(* Logix 5000 project; controller TFF vendor 1 type 14 code 107 rev 33.11; software revision 33.04; part 17 of 38 *)
(* tags used below, declared in another part *)
   PCV101_AutoMaxRate : REAL;   // PCV101 Maximum Rate in Auto Mode
   PCV101_ManualMaxRate : REAL;   // PCV101 Maximum Rate in Manual mode
   PCV101_Max_CV : REAL;   // Max CV for PCV101
   ControlLoop : ControlLoop[20];   // Control Loop Array
   ControlLoop_PCV101 : ALIAS FOR ControlLoop[3];
   ControlLoop_PCV101_5ms : ALIAS FOR ControlLoop[4];
   ControlLoop_PCV101Alarm : ALIAS FOR AlarmDeviation[3];
   ControlLoop_PCV201 : ALIAS FOR ControlLoop[5];
   ControlLoop_PCV201_5ms : ALIAS FOR ControlLoop[6];
   ControlLoop_PCV201_RAMP_OUT : REAL;   // Ramp Output
   PCV101 : ALIAS FOR AnalogPoint[3];
   PCV101_AO : ALIAS FOR AnalogOutput[3];
   PCV101_Control : PCV_Control;   // PCV101 Control UDT
   PCV101_CVTune : CVTune;
   PCV101_PID : PCV;   // PCV101 PID Management
   PCV201 : ALIAS FOR AnalogPoint[4];
   PCV201_Control : PCV_Control;   // PCV201 Control UDT
   PCV201_PID : PCV;   // PCV201 PID Management
   Rack_Murr_Node1_TFF20 : IO_Station;   // Status of Node 1 TFF20
   Rack_Murr_Node1_TFF40 : IO_Station;   // Status of Node 1 TFF40
   Rack_Murr_Node1_TFF80 : IO_Station;   // Status of Node 1 TFF80
   RawAnalogInputArray : INT[50];   // Array of analog input raw
   SysControl : SysControl;   // General system status and command
   ThisSystem : SystemType;
   TMP : ALIAS FOR AnalogPoint[41];
   Valve : Valve[100];   // Valve Array
(* MainProgram5ms, continued *)

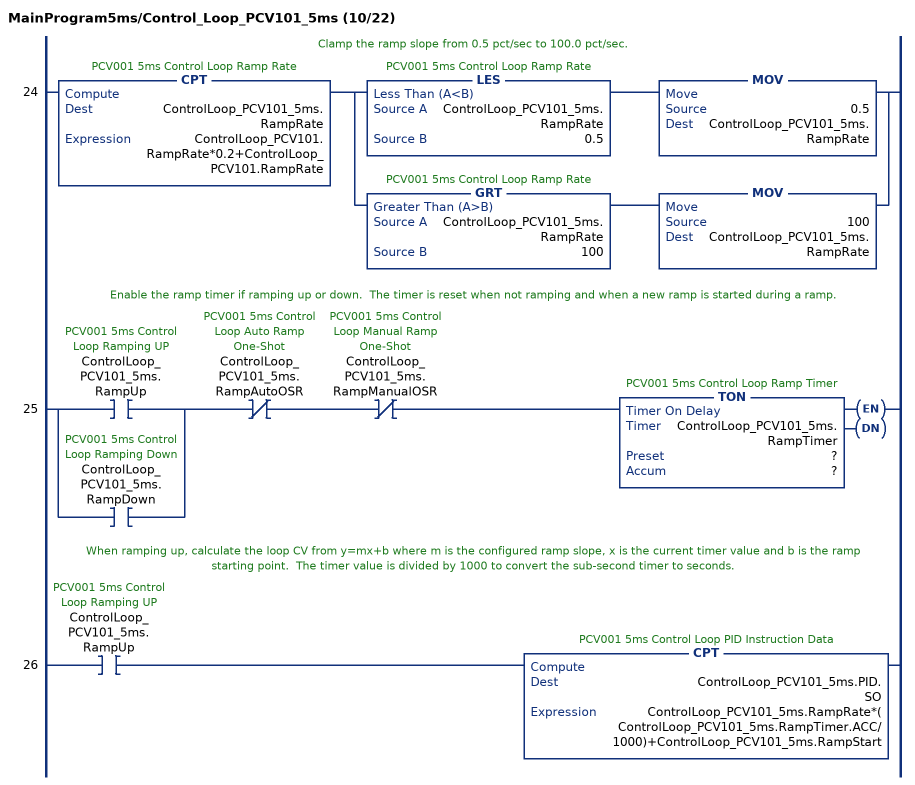
   [picture p62: MainProgram5ms/Control_Loop_PCV101_5ms rungs 24-26]
   // Clamp the ramp slope from 0.5 pct/sec to 100.0 pct/sec.
   24: CPT(ControlLoop_PCV101_5ms.RampRate,ControlLoop_PCV101.RampRate*0.2+ControlLoop_PCV101.RampRate)[LES(ControlLoop_PCV101_5ms.RampRate,0.5) MOV(0.5,ControlLoop_PCV101_5ms.RampRate) ,GRT(ControlLoop_PCV101_5ms.RampRate,100) MOV(100,ControlLoop_PCV101_5ms.RampRate) ];
   // Enable the ramp timer if ramping up or down.  The timer is reset when not ramping and when a new ramp is started during a ramp.
   25: [XIC(ControlLoop_PCV101_5ms.RampUp) ,XIC(ControlLoop_PCV101_5ms.RampDown) ]XIO(ControlLoop_PCV101_5ms.RampAutoOSR)XIO(ControlLoop_PCV101_5ms.RampManualOSR)TON(ControlLoop_PCV101_5ms.RampTimer,?,?);
   // When ramping up, calculate the loop CV from y=mx+b where m is the configured ramp slope, x is the current timer value and b is the ramp starting point.  The timer value is divided by 1000 to convert the sub-second timer to seconds.
   26: XIC(ControlLoop_PCV101_5ms.RampUp)CPT(ControlLoop_PCV101_5ms.PID.SO,ControlLoop_PCV101_5ms.RampRate*(ControlLoop_PCV101_5ms.RampTimer.ACC/1000)+ControlLoop_PCV101_5ms.RampStart);
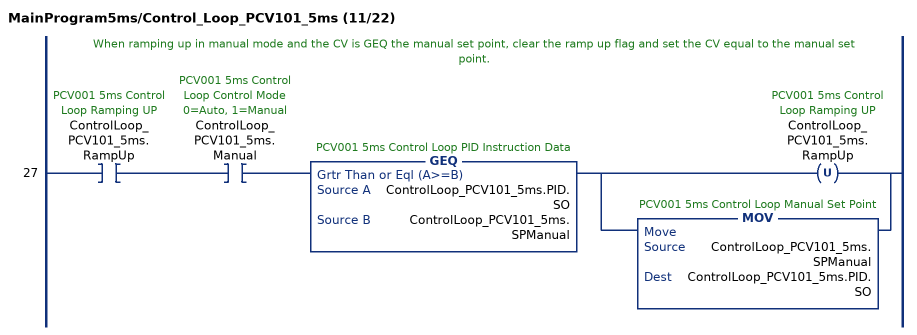
   // When ramping up in manual mode and the CV is GEQ the manual set point, clear the ramp up flag and set the CV equal to the manual set point.
   27: XIC(ControlLoop_PCV101_5ms.RampUp)XIC(ControlLoop_PCV101_5ms.Manual)GEQ(ControlLoop_PCV101_5ms.PID.SO,ControlLoop_PCV101_5ms.SPManual)[OTU(ControlLoop_PCV101_5ms.RampUp) ,MOV(ControlLoop_PCV101_5ms.SPManual,ControlLoop_PCV101_5ms.PID.SO) ];
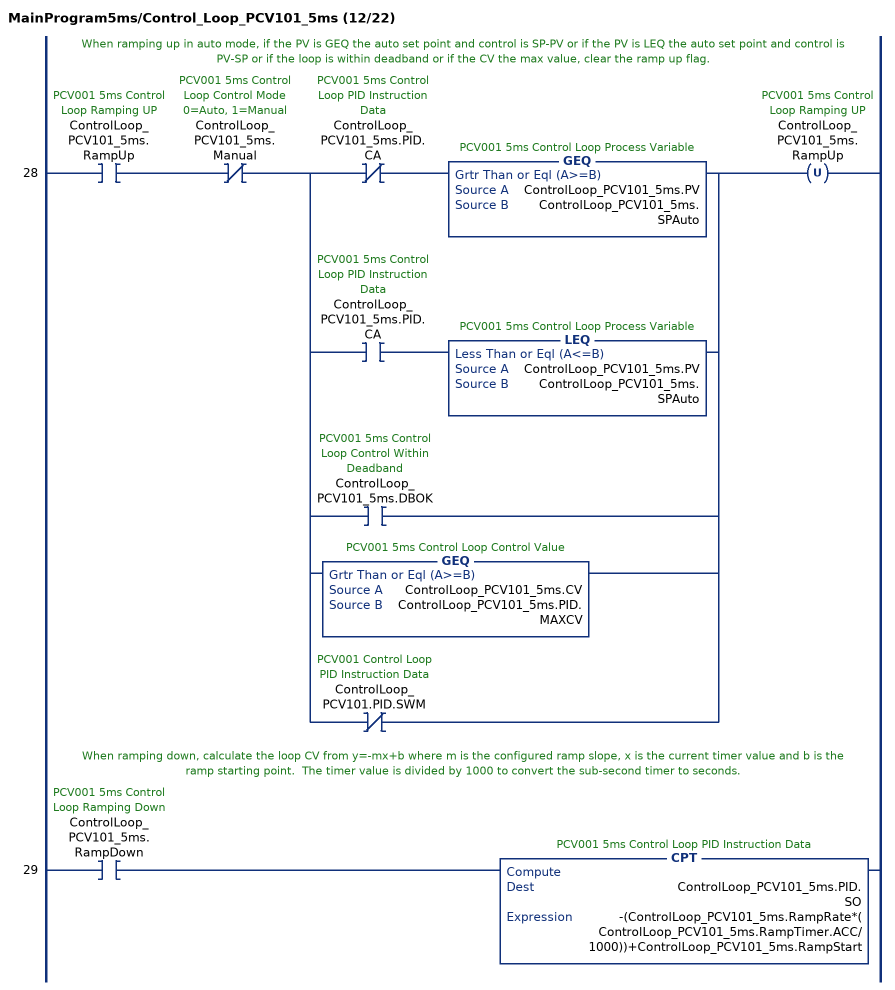
   // When ramping up in auto mode, if the PV is GEQ the auto set point and control is SP-PV or if the PV is LEQ the auto set point and control is PV-SP or if the loop is within deadband or if the CV the max value, clear the ramp up flag.
   28: XIC(ControlLoop_PCV101_5ms.RampUp)XIO(ControlLoop_PCV101_5ms.Manual)[XIO(ControlLoop_PCV101_5ms.PID.CA) GEQ(ControlLoop_PCV101_5ms.PV,ControlLoop_PCV101_5ms.SPAuto) ,XIC(ControlLoop_PCV101_5ms.PID.CA) LEQ(ControlLoop_PCV101_5ms.PV,ControlLoop_PCV101_5ms.SPAuto) ,XIC(ControlLoop_PCV101_5ms.DBOK) ,[GEQ(ControlLoop_PCV101_5ms.CV,ControlLoop_PCV101_5ms.PID.MAXCV) ,XIO(ControlLoop_PCV101.PID.SWM) ] ]OTU(ControlLoop_PCV101_5ms.RampUp);
   // When ramping down, calculate the loop CV from y=-mx+b where m is the configured ramp slope, x is the current timer value and b is the ramp starting point.  The timer value is divided by 1000 to convert the sub-second timer to seconds.
   29: XIC(ControlLoop_PCV101_5ms.RampDown)CPT(ControlLoop_PCV101_5ms.PID.SO,-(ControlLoop_PCV101_5ms.RampRate*(ControlLoop_PCV101_5ms.RampTimer.ACC/1000))+ControlLoop_PCV101_5ms.RampStart);
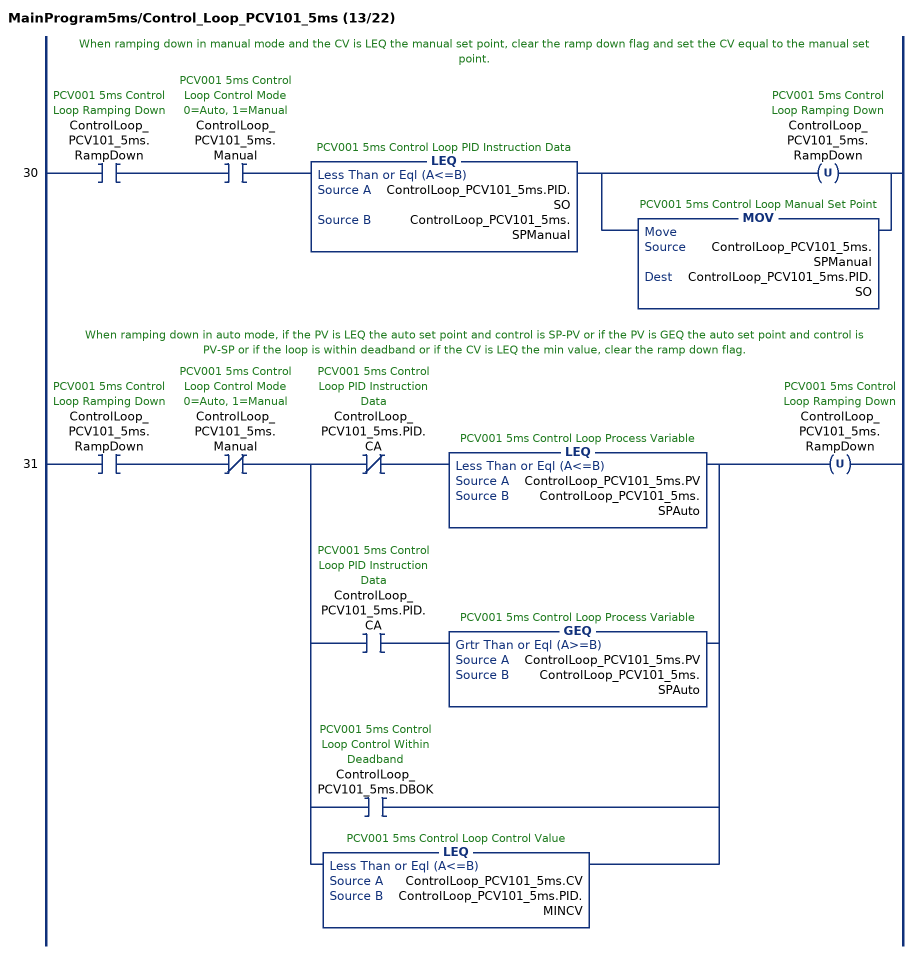
   // When ramping down in manual mode and the CV is LEQ the manual set point, clear the ramp down flag and set the CV equal to the manual set point.
   30: XIC(ControlLoop_PCV101_5ms.RampDown)XIC(ControlLoop_PCV101_5ms.Manual)LEQ(ControlLoop_PCV101_5ms.PID.SO,ControlLoop_PCV101_5ms.SPManual)[OTU(ControlLoop_PCV101_5ms.RampDown) ,MOV(ControlLoop_PCV101_5ms.SPManual,ControlLoop_PCV101_5ms.PID.SO) ];
   // When ramping down in auto mode, if the PV is LEQ the auto set point and control is SP-PV or if the PV is GEQ the auto set point and control is PV-SP or if the loop is within deadband or if the CV is LEQ the min value, clear the ramp down flag.
   31: XIC(ControlLoop_PCV101_5ms.RampDown)XIO(ControlLoop_PCV101_5ms.Manual)[XIO(ControlLoop_PCV101_5ms.PID.CA) LEQ(ControlLoop_PCV101_5ms.PV,ControlLoop_PCV101_5ms.SPAuto) ,XIC(ControlLoop_PCV101_5ms.PID.CA) GEQ(ControlLoop_PCV101_5ms.PV,ControlLoop_PCV101_5ms.SPAuto) ,XIC(ControlLoop_PCV101_5ms.DBOK) ,LEQ(ControlLoop_PCV101_5ms.CV,ControlLoop_PCV101_5ms.PID.MINCV) ]OTU(ControlLoop_PCV101_5ms.RampDown);
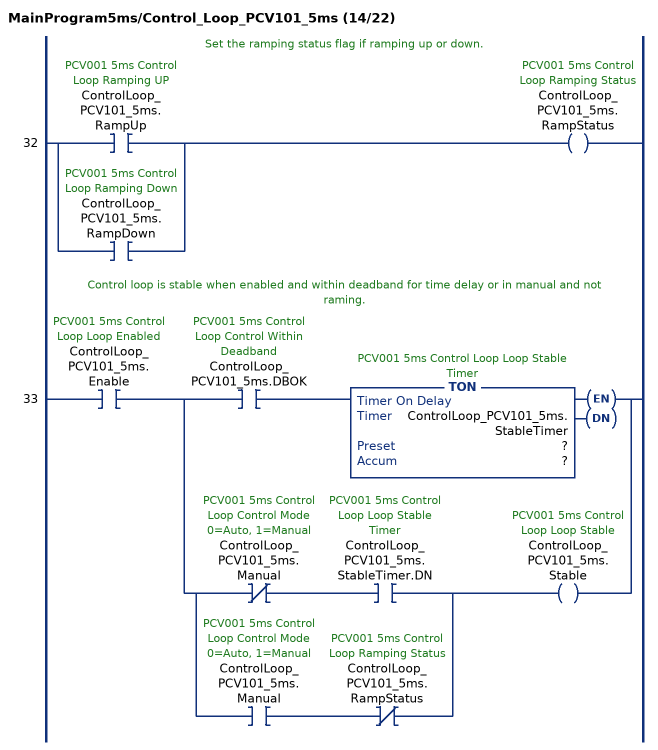
   // Set the ramping status flag if ramping up or down.
   32: [XIC(ControlLoop_PCV101_5ms.RampUp) ,XIC(ControlLoop_PCV101_5ms.RampDown) ]OTE(ControlLoop_PCV101_5ms.RampStatus);
   // Control loop is stable when enabled and within deadband for time delay or in manual and not raming.
   33: XIC(ControlLoop_PCV101_5ms.Enable)[XIC(ControlLoop_PCV101_5ms.DBOK) TON(ControlLoop_PCV101_5ms.StableTimer,?,?) ,[XIO(ControlLoop_PCV101_5ms.Manual) XIC(ControlLoop_PCV101_5ms.StableTimer.DN) ,XIC(ControlLoop_PCV101_5ms.Manual) XIO(ControlLoop_PCV101_5ms.RampStatus) ] OTE(ControlLoop_PCV101_5ms.Stable) ];
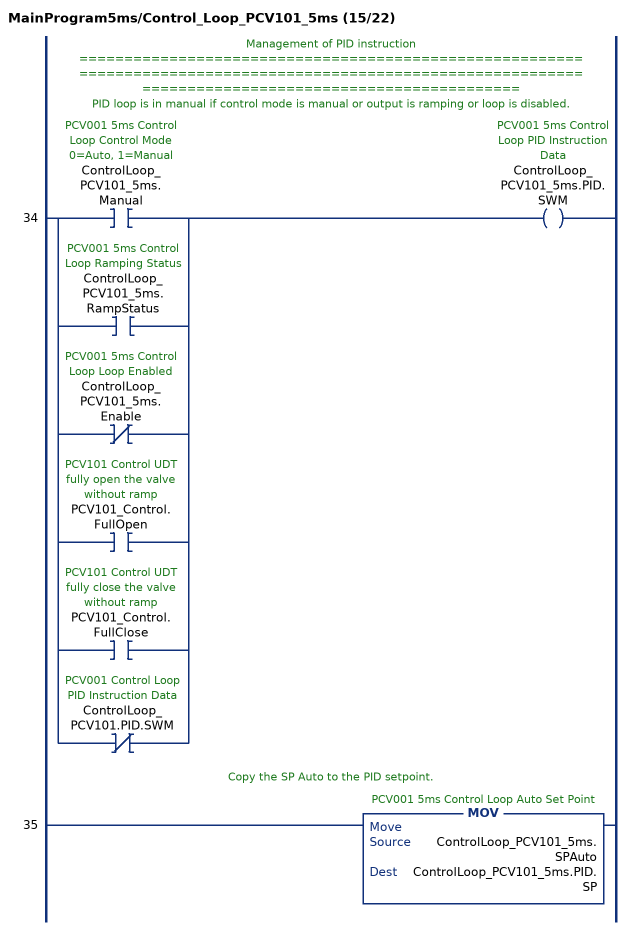
   // Management of PID instruction
   // ==========================================================================================================================================================
   // PID loop is in manual if control mode is manual or output is ramping or loop is disabled.
   34: [XIC(ControlLoop_PCV101_5ms.Manual) ,XIC(ControlLoop_PCV101_5ms.RampStatus) ,XIO(ControlLoop_PCV101_5ms.Enable) ,[[XIC(PCV101_Control.FullOpen) ,XIC(PCV101_Control.FullClose) ] ,XIO(ControlLoop_PCV101.PID.SWM) ] ]OTE(ControlLoop_PCV101_5ms.PID.SWM);
   // Copy the SP Auto to the PID setpoint.
   35: MOV(ControlLoop_PCV101_5ms.SPAuto,ControlLoop_PCV101_5ms.PID.SP);
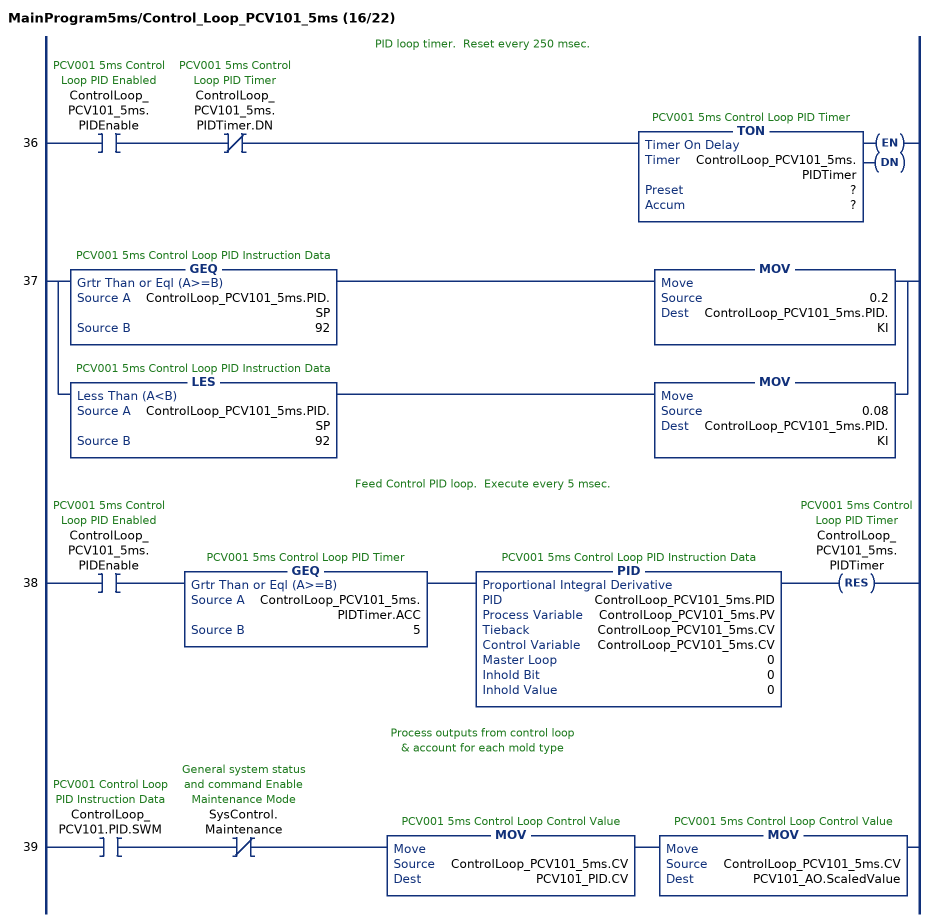
   // PID loop timer.  Reset every 250 msec.
   36: XIC(ControlLoop_PCV101_5ms.PIDEnable)XIO(ControlLoop_PCV101_5ms.PIDTimer.DN)TON(ControlLoop_PCV101_5ms.PIDTimer,?,?);
   37: [GEQ(ControlLoop_PCV101_5ms.PID.SP,92) MOV(0.2,ControlLoop_PCV101_5ms.PID.KI) ,LES(ControlLoop_PCV101_5ms.PID.SP,92) MOV(0.08,ControlLoop_PCV101_5ms.PID.KI) ];
   // Feed Control PID loop.  Execute every 5 msec.
   38: XIC(ControlLoop_PCV101_5ms.PIDEnable)GEQ(ControlLoop_PCV101_5ms.PIDTimer.ACC,5)PID(ControlLoop_PCV101_5ms.PID,ControlLoop_PCV101_5ms.PV,ControlLoop_PCV101_5ms.CV,ControlLoop_PCV101_5ms.CV,0,0,0)RES(ControlLoop_PCV101_5ms.PIDTimer);
   // Process outputs from control loop
   // & account for each mold type
   39: XIC(ControlLoop_PCV101.PID.SWM)XIO(SysControl.Maintenance)MOV(ControlLoop_PCV101_5ms.CV,PCV101_PID.CV)MOV(ControlLoop_PCV101_5ms.CV,PCV101_AO.ScaledValue);
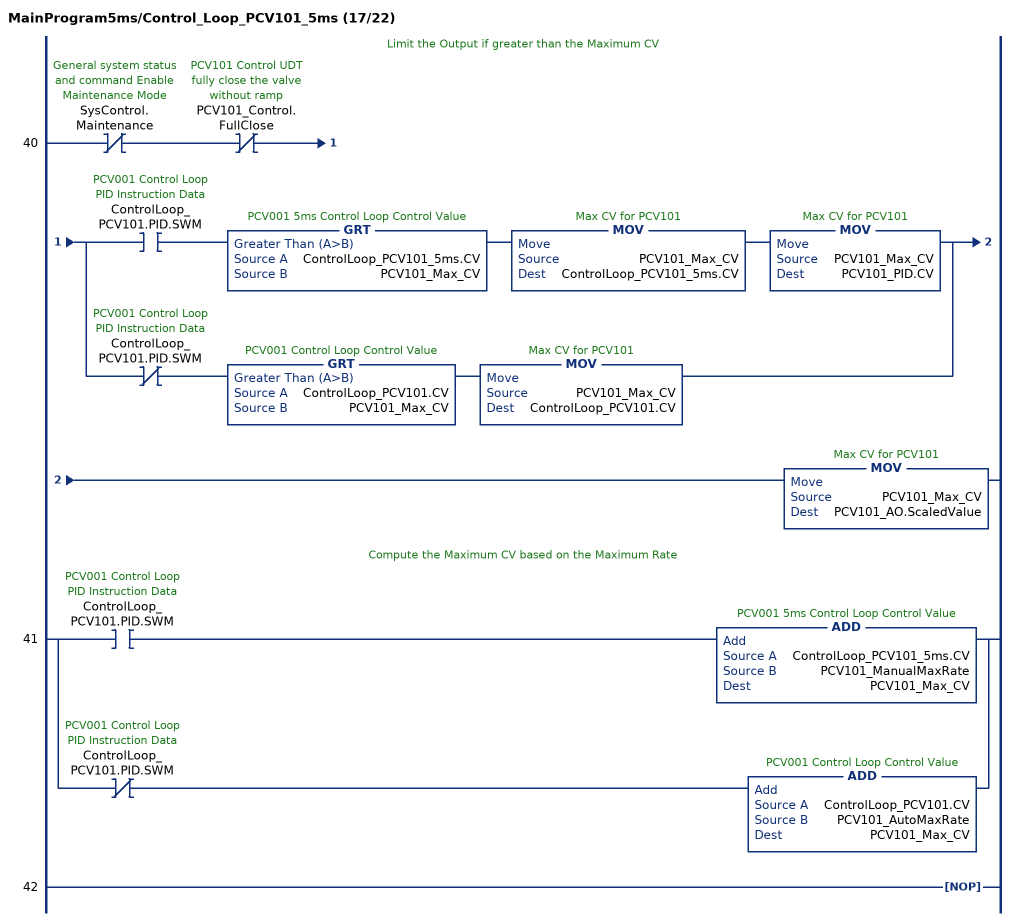
   // Limit the Output if greater than the Maximum CV
   40: XIO(SysControl.Maintenance)XIO(PCV101_Control.FullClose)[XIC(ControlLoop_PCV101.PID.SWM) GRT(ControlLoop_PCV101_5ms.CV,PCV101_Max_CV) MOV(PCV101_Max_CV,ControlLoop_PCV101_5ms.CV) MOV(PCV101_Max_CV,PCV101_PID.CV) ,XIO(ControlLoop_PCV101.PID.SWM) GRT(ControlLoop_PCV101.CV,PCV101_Max_CV) MOV(PCV101_Max_CV,ControlLoop_PCV101.CV) ]MOV(PCV101_Max_CV,PCV101_AO.ScaledValue);
   // Compute the Maximum CV based on the Maximum Rate
   41: [XIC(ControlLoop_PCV101.PID.SWM) ADD(ControlLoop_PCV101_5ms.CV,PCV101_ManualMaxRate,PCV101_Max_CV) ,XIO(ControlLoop_PCV101.PID.SWM) ADD(ControlLoop_PCV101.CV,PCV101_AutoMaxRate,PCV101_Max_CV) ];
   42: NOP();
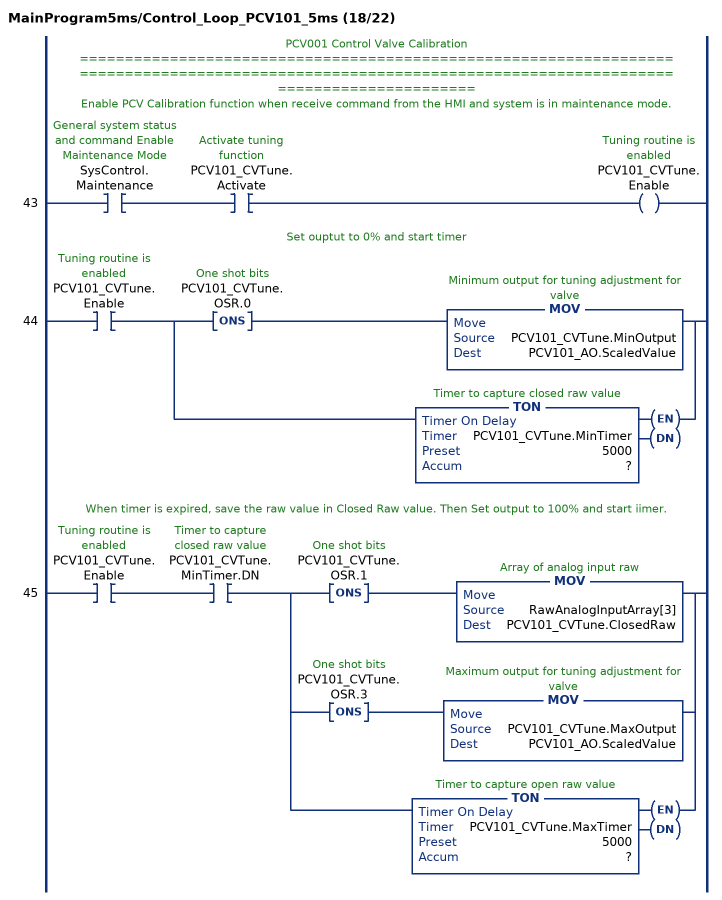
   // PCV001 Control Valve Calibration
   // ==========================================================================================================================================================
   // Enable PCV Calibration function when receive command from the HMI and system is in maintenance mode.
   43: XIC(SysControl.Maintenance)XIC(PCV101_CVTune.Activate)OTE(PCV101_CVTune.Enable);
   // Set ouptut to 0% and start timer
   44: XIC(PCV101_CVTune.Enable)[ONS(PCV101_CVTune.OSR.0) MOV(PCV101_CVTune.MinOutput,PCV101_AO.ScaledValue) ,TON(PCV101_CVTune.MinTimer,?,?) ];
   // When timer is expired, save the raw value in Closed Raw value. Then Set output to 100% and start iimer.
   45: XIC(PCV101_CVTune.Enable)XIC(PCV101_CVTune.MinTimer.DN)[ONS(PCV101_CVTune.OSR.1) MOV(RawAnalogInputArray[3],PCV101_CVTune.ClosedRaw) ,ONS(PCV101_CVTune.OSR.3) MOV(PCV101_CVTune.MaxOutput,PCV101_AO.ScaledValue) ,TON(PCV101_CVTune.MaxTimer,?,?) ];
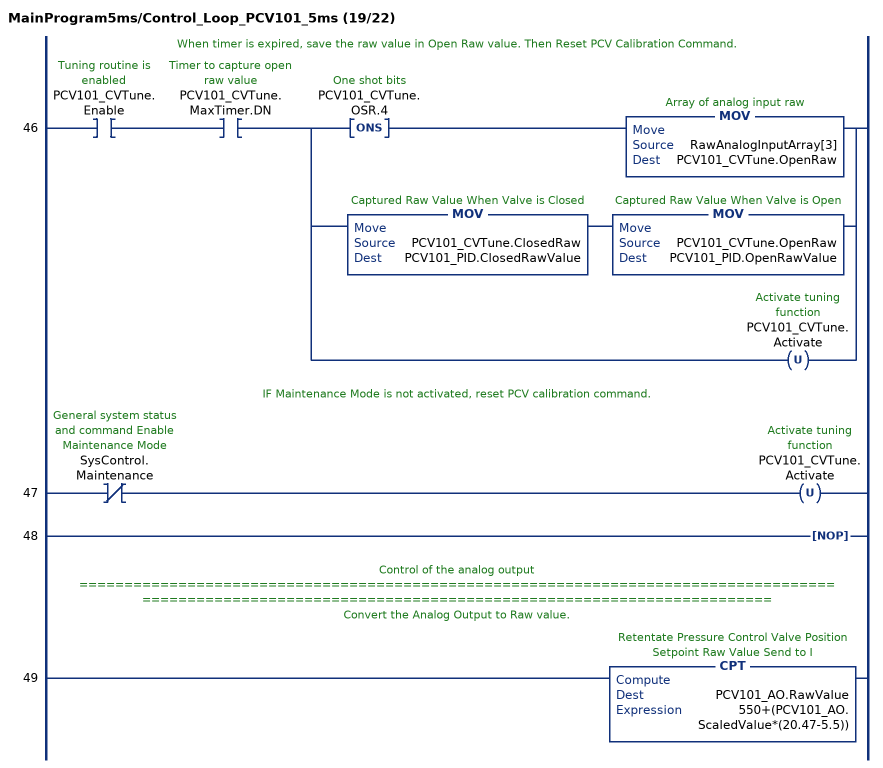
   // When timer is expired, save the raw value in Open Raw value. Then Reset PCV Calibration Command.
   46: XIC(PCV101_CVTune.Enable)XIC(PCV101_CVTune.MaxTimer.DN)[ONS(PCV101_CVTune.OSR.4) MOV(RawAnalogInputArray[3],PCV101_CVTune.OpenRaw) ,MOV(PCV101_CVTune.ClosedRaw,PCV101_PID.ClosedRawValue) MOV(PCV101_CVTune.OpenRaw,PCV101_PID.OpenRawValue) ,OTU(PCV101_CVTune.Activate) ];
   // IF Maintenance Mode is not activated, reset PCV calibration command.
   47: XIO(SysControl.Maintenance)OTU(PCV101_CVTune.Activate);
   48: NOP();
   // Control of the analog output
   // ==========================================================================================================================================================
   // Convert the Analog Output to Raw value.
   49: CPT(PCV101_AO.RawValue,550+(PCV101_AO.ScaledValue*(20.47-5.5)));
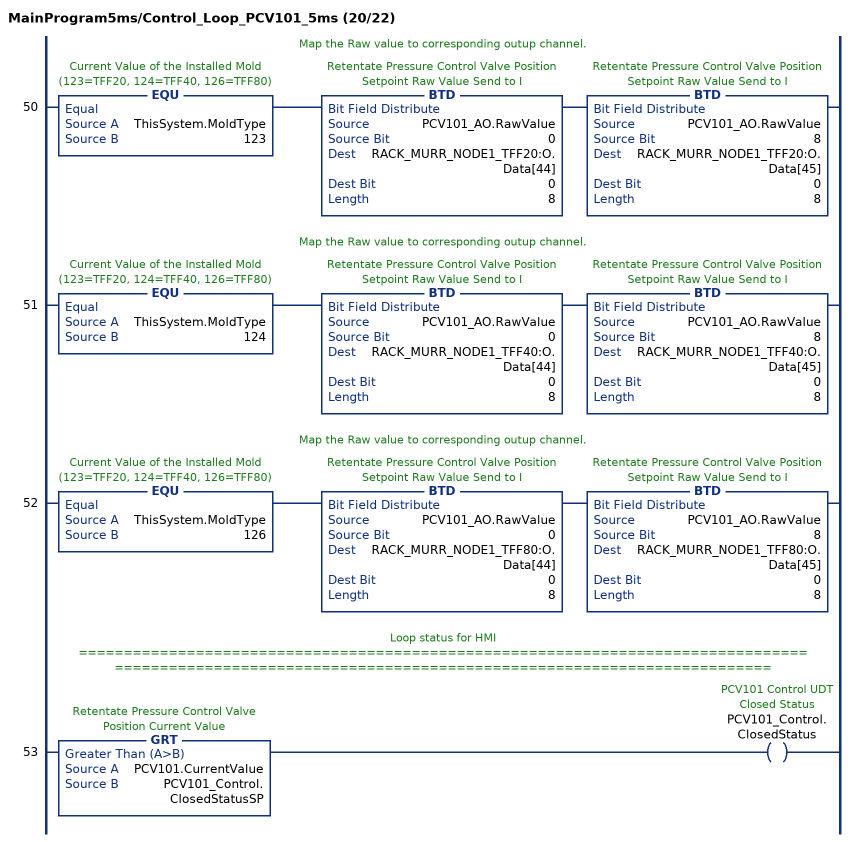
   // Map the Raw value to corresponding outup channel.
   50: EQU(ThisSystem.MoldType,123)BTD(PCV101_AO.RawValue,0,RACK_MURR_NODE1_TFF20:O.Data[44],0,8)BTD(PCV101_AO.RawValue,8,RACK_MURR_NODE1_TFF20:O.Data[45],0,8);
   // Map the Raw value to corresponding outup channel.
   51: EQU(ThisSystem.MoldType,124)BTD(PCV101_AO.RawValue,0,RACK_MURR_NODE1_TFF40:O.Data[44],0,8)BTD(PCV101_AO.RawValue,8,RACK_MURR_NODE1_TFF40:O.Data[45],0,8);
   // Map the Raw value to corresponding outup channel.
   52: EQU(ThisSystem.MoldType,126)BTD(PCV101_AO.RawValue,0,RACK_MURR_NODE1_TFF80:O.Data[44],0,8)BTD(PCV101_AO.RawValue,8,RACK_MURR_NODE1_TFF80:O.Data[45],0,8);
   // Loop status for HMI
   // ==========================================================================================================================================================
   53: GRT(PCV101.CurrentValue,PCV101_Control.ClosedStatusSP)OTE(PCV101_Control.ClosedStatus);
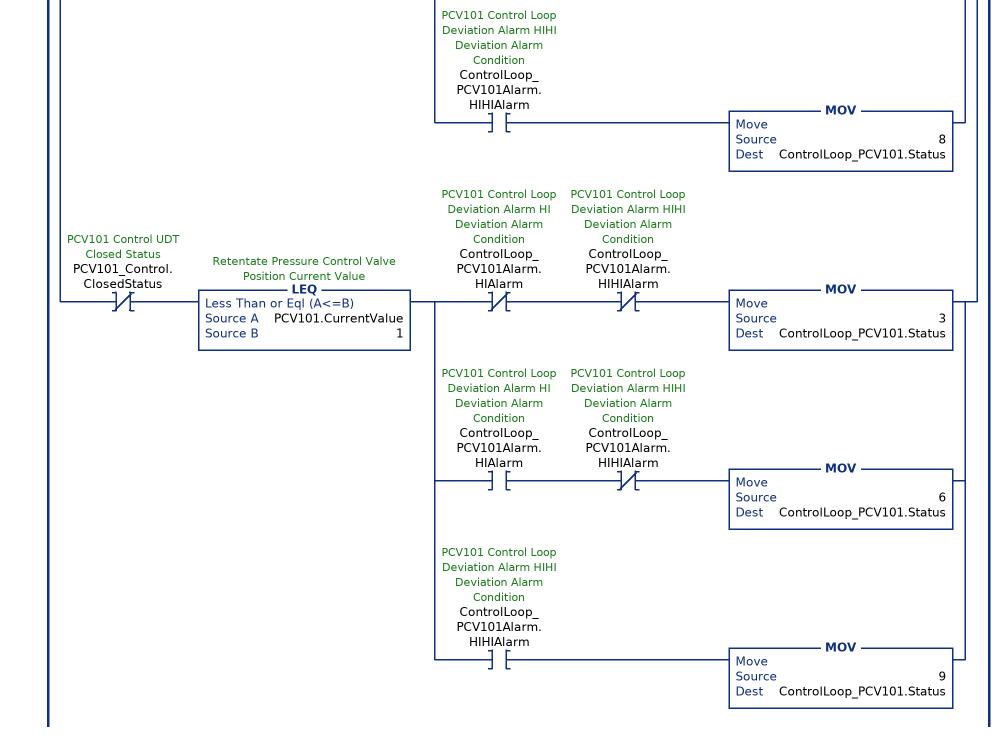
   // ControlLoop Status : 1 = PCV Close
   // ControlLoop Status : 2 = PCV Open
   // ControlLoop Status : 3 = PCV Full Open
   // ControlLoop Status : 4 = PCV Close and Non Critical alam
   // ControlLoop Status : 5 = PCV Open and Non Critical alam
   // ControlLoop Status : 6 = PCV Full Open and Non Critical alam
   // ControlLoop Status : 7 = PCV Close and Critical alam
   // ControlLoop Status : 8 = PCV Open and Critical alam
   // ControlLoop Status : 9 = PCV Full Open and Critical alam
   54: [XIC(PCV101_Control.ClosedStatus) [XIO(ControlLoop_PCV101Alarm.HIAlarm) XIO(ControlLoop_PCV101Alarm.HIHIAlarm) MOV(1,ControlLoop_PCV101.Status) ,XIC(ControlLoop_PCV101Alarm.HIAlarm) XIO(ControlLoop_PCV101Alarm.HIHIAlarm) MOV(4,ControlLoop_PCV101.Status) ,XIC(ControlLoop_PCV101Alarm.HIHIAlarm) MOV(7,ControlLoop_PCV101.Status) ] ,XIO(PCV101_Control.ClosedStatus) GRT(PCV101.CurrentValue,2) [XIO(ControlLoop_PCV101Alarm.HIAlarm) XIO(ControlLoop_PCV101Alarm.HIHIAlarm) MOV(2,ControlLoop_PCV101.Status) ,XIC(ControlLoop_PCV101Alarm.HIAlarm) XIO(ControlLoop_PCV101Alarm.HIHIAlarm) MOV(5,ControlLoop_PCV101.Status) ,XIC(ControlLoop_PCV101Alarm.HIHIAlarm) MOV(8,ControlLoop_PCV101.Status) ] ,XIO(PCV101_Control.ClosedStatus) LEQ(PCV101.CurrentValue,1) [XIO(ControlLoop_PCV101Alarm.HIAlarm) XIO(ControlLoop_PCV101Alarm.HIHIAlarm) MOV(3,ControlLoop_PCV101.Status) ,XIC(ControlLoop_PCV101Alarm.HIAlarm) XIO(ControlLoop_PCV101Alarm.HIHIAlarm) MOV(6,ControlLoop_PCV101.Status) ,XIC(ControlLoop_PCV101Alarm.HIHIAlarm) MOV(9,ControlLoop_PCV101.Status) ] ];
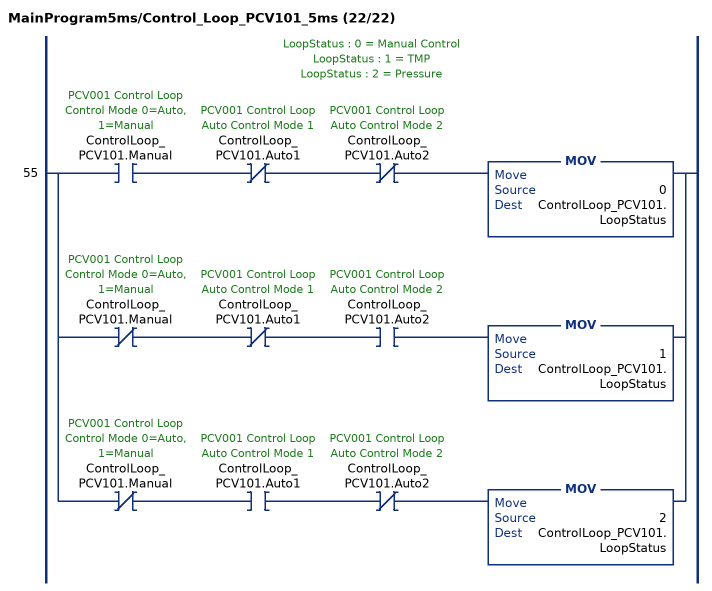
   // LoopStatus : 0 = Manual Control
   //  LoopStatus : 1 = TMP
   //  LoopStatus : 2 = Pressure
   55: [XIC(ControlLoop_PCV101.Manual) XIO(ControlLoop_PCV101.Auto1) XIO(ControlLoop_PCV101.Auto2) MOV(0,ControlLoop_PCV101.LoopStatus) ,XIO(ControlLoop_PCV101.Manual) XIO(ControlLoop_PCV101.Auto1) XIC(ControlLoop_PCV101.Auto2) MOV(1,ControlLoop_PCV101.LoopStatus) ,XIO(ControlLoop_PCV101.Manual) XIC(ControlLoop_PCV101.Auto1) XIO(ControlLoop_PCV101.Auto2) MOV(2,ControlLoop_PCV101.LoopStatus) ];
END_ROUTINE

ROUTINE Control_Loop_PCV201_5ms   (* ladder *)
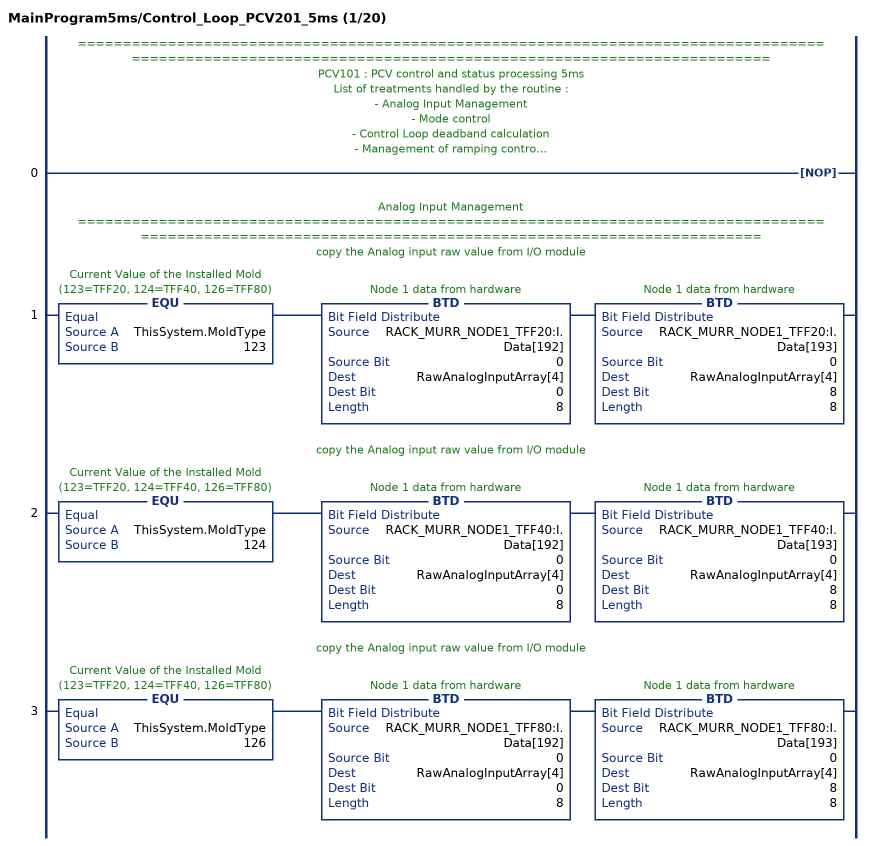
   // ==========================================================================================================================================================
   //                                                  PCV101 : PCV control and status processing 5ms
   //                                                     List of treatments handled by the routine :
   //                                                           - Analog Input Management
   //                                                          - Mode control
   //                                                          - Control Loop deadband calculation
   //                                                          - Management of ramping control
   //                                                          - Management of PID instruction
   //                                                          - PCV101 Control Valve Calibration
   //                                                          - Control of the analog output
   //                                                          - Loop status for HMI
   //                                                     -----------------------------------------------------------------------------------------------------------------------------------------------------
   //                                                     History
   // 		2019-DEC-24 - Merck - Q. Spindler - Initial version for Candidate Release 1.00.00.00.a
   // 		2021-APR-19 - Merck - Q. Spindler - Modifications for Candidate Release 1.00.00.00.e
   //                                                    - Start the PCV to close at 550 point instead of 0 (a bit less than 2 bar)
   // ==========================================================================================================================================================
   0: NOP();
   // Analog Input Management
   // ========================================================================================================================================================
   // copy the Analog input raw value from I/O module
   1: EQU(ThisSystem.MoldType,123)BTD(RACK_MURR_NODE1_TFF20:I.Data[192],0,RawAnalogInputArray[4],0,8)BTD(RACK_MURR_NODE1_TFF20:I.Data[193],0,RawAnalogInputArray[4],8,8);
   // copy the Analog input raw value from I/O module
   2: EQU(ThisSystem.MoldType,124)BTD(RACK_MURR_NODE1_TFF40:I.Data[192],0,RawAnalogInputArray[4],0,8)BTD(RACK_MURR_NODE1_TFF40:I.Data[193],0,RawAnalogInputArray[4],8,8);
   // copy the Analog input raw value from I/O module
   3: EQU(ThisSystem.MoldType,126)BTD(RACK_MURR_NODE1_TFF80:I.Data[192],0,RawAnalogInputArray[4],0,8)BTD(RACK_MURR_NODE1_TFF80:I.Data[193],0,RawAnalogInputArray[4],8,8);
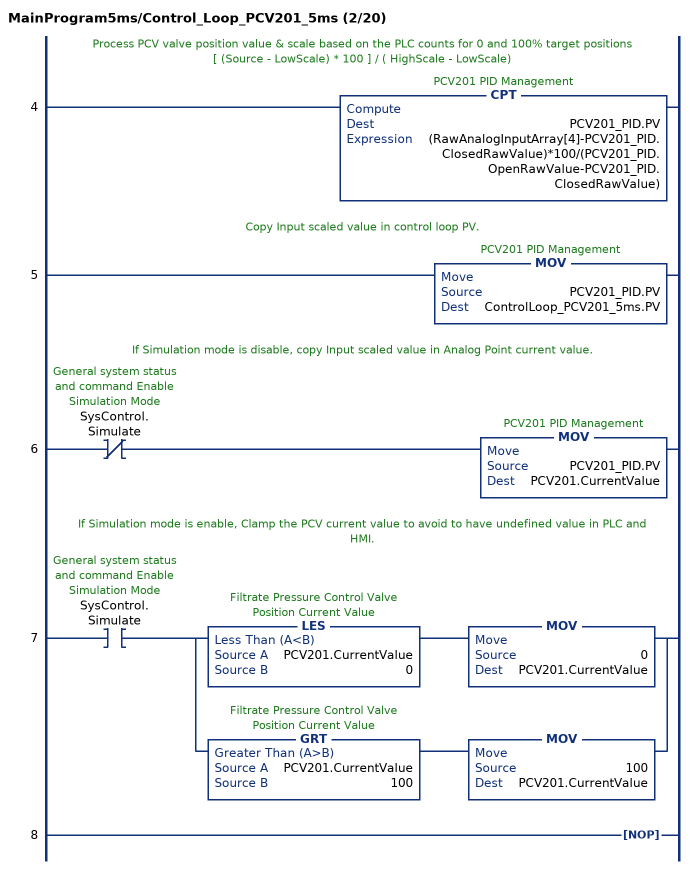
   // Process PCV valve position value & scale based on the PLC counts for 0 and 100% target positions
   // [ (Source - LowScale) * 100 ] / ( HighScale - LowScale)
   4: CPT(PCV201_PID.PV,(RawAnalogInputArray[4]-PCV201_PID.ClosedRawValue)*100/(PCV201_PID.OpenRawValue-PCV201_PID.ClosedRawValue));
   // Copy Input scaled value in control loop PV.
   5: MOV(PCV201_PID.PV,ControlLoop_PCV201_5ms.PV);
   // If Simulation mode is disable, copy Input scaled value in Analog Point current value.
   6: XIO(SysControl.Simulate)MOV(PCV201_PID.PV,PCV201.CurrentValue);
   // If Simulation mode is enable, Clamp the PCV current value to avoid to have undefined value in PLC and HMI.
   7: XIC(SysControl.Simulate)[LES(PCV201.CurrentValue,0) MOV(0,PCV201.CurrentValue) ,GRT(PCV201.CurrentValue,100) MOV(100,PCV201.CurrentValue) ];
   8: NOP();
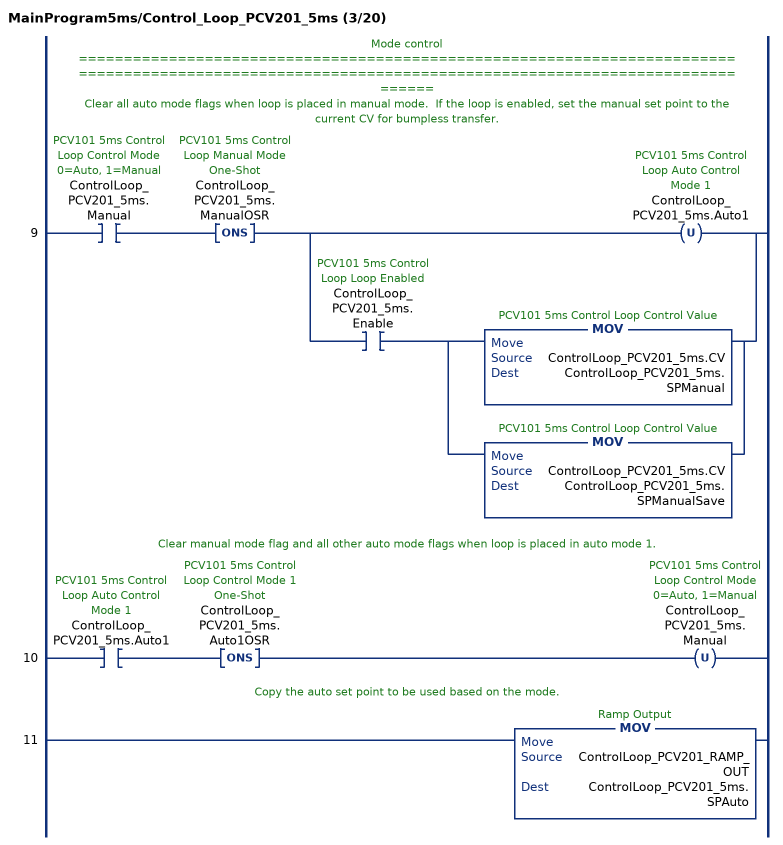
   // Mode control
   // ========================================================================================================================================================
   // Clear all auto mode flags when loop is placed in manual mode.  If the loop is enabled, set the manual set point to the current CV for bumpless transfer.
   9: XIC(ControlLoop_PCV201_5ms.Manual)ONS(ControlLoop_PCV201_5ms.ManualOSR)[OTU(ControlLoop_PCV201_5ms.Auto1) ,XIC(ControlLoop_PCV201_5ms.Enable) [MOV(ControlLoop_PCV201_5ms.CV,ControlLoop_PCV201_5ms.SPManual) ,MOV(ControlLoop_PCV201_5ms.CV,ControlLoop_PCV201_5ms.SPManualSave) ] ];
   // Clear manual mode flag and all other auto mode flags when loop is placed in auto mode 1.
   10: XIC(ControlLoop_PCV201_5ms.Auto1)ONS(ControlLoop_PCV201_5ms.Auto1OSR)OTU(ControlLoop_PCV201_5ms.Manual);
   // Copy the auto set point to be used based on the mode.
   11: MOV(ControlLoop_PCV201_RAMP_OUT,ControlLoop_PCV201_5ms.SPAuto);
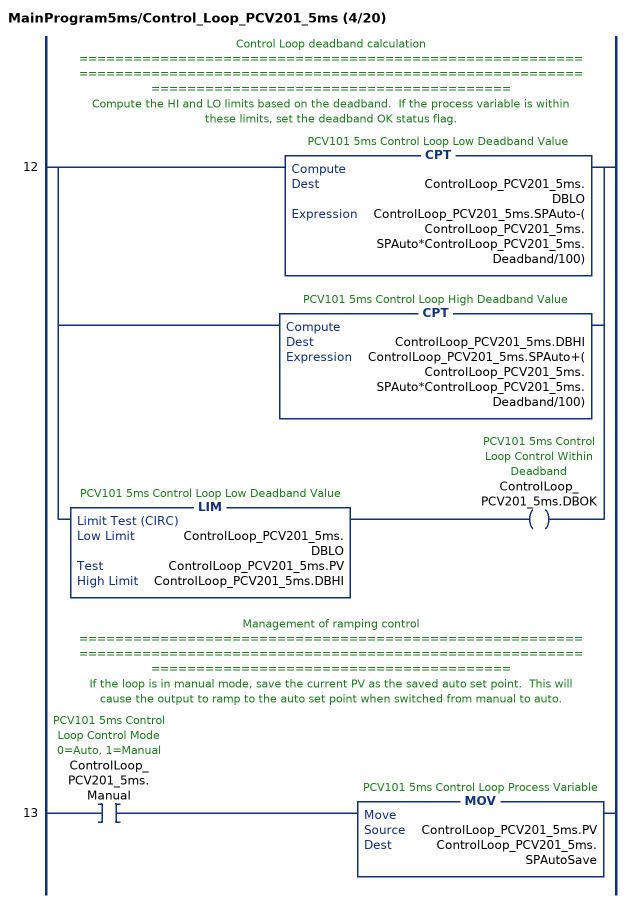
   // Control Loop deadband calculation
   // ========================================================================================================================================================
   // Compute the HI and LO limits based on the deadband.  If the process variable is within these limits, set the deadband OK status flag.
   12: [CPT(ControlLoop_PCV201_5ms.DBLO,ControlLoop_PCV201_5ms.SPAuto-(ControlLoop_PCV201_5ms.SPAuto*ControlLoop_PCV201_5ms.Deadband/100)) ,CPT(ControlLoop_PCV201_5ms.DBHI,ControlLoop_PCV201_5ms.SPAuto+(ControlLoop_PCV201_5ms.SPAuto*ControlLoop_PCV201_5ms.Deadband/100)) ,LIM(ControlLoop_PCV201_5ms.DBLO,ControlLoop_PCV201_5ms.PV,ControlLoop_PCV201_5ms.DBHI) OTE(ControlLoop_PCV201_5ms.DBOK) ];
   // Management of ramping control
   // ========================================================================================================================================================
   // If the loop is in manual mode, save the current PV as the saved auto set point.  This will cause the output to ramp to the auto set point when switched from manual to auto.
   13: XIC(ControlLoop_PCV201_5ms.Manual)MOV(ControlLoop_PCV201_5ms.PV,ControlLoop_PCV201_5ms.SPAutoSave);
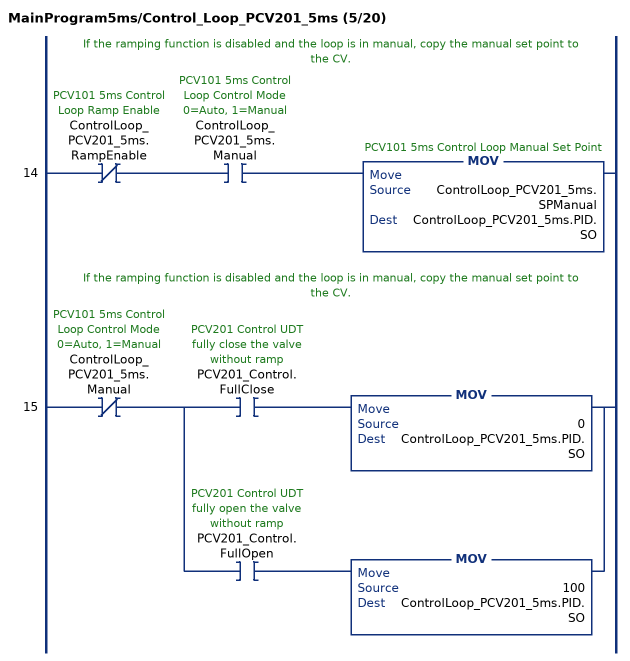
   // If the ramping function is disabled and the loop is in manual, copy the manual set point to the CV.
   14: XIO(ControlLoop_PCV201_5ms.RampEnable)XIC(ControlLoop_PCV201_5ms.Manual)MOV(ControlLoop_PCV201_5ms.SPManual,ControlLoop_PCV201_5ms.PID.SO);
   // If the ramping function is disabled and the loop is in manual, copy the manual set point to the CV.
   15: XIO(ControlLoop_PCV201_5ms.Manual)[XIC(PCV201_Control.FullClose) MOV(0,ControlLoop_PCV201_5ms.PID.SO) ,XIC(PCV201_Control.FullOpen) MOV(100,ControlLoop_PCV201_5ms.PID.SO) ];
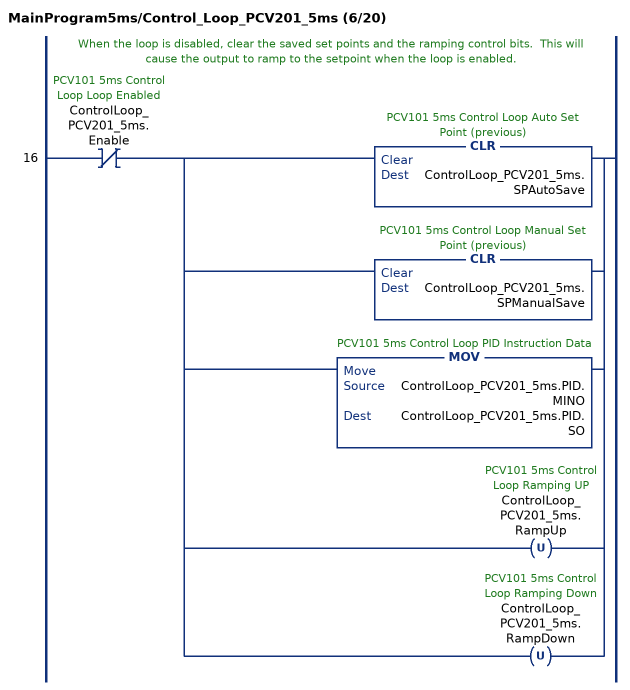
   // When the loop is disabled, clear the saved set points and the ramping control bits.  This will cause the output to ramp to the setpoint when the loop is enabled.
   16: XIO(ControlLoop_PCV201_5ms.Enable)[CLR(ControlLoop_PCV201_5ms.SPAutoSave) ,CLR(ControlLoop_PCV201_5ms.SPManualSave) ,MOV(ControlLoop_PCV201_5ms.PID.MINO,ControlLoop_PCV201_5ms.PID.SO) ,OTU(ControlLoop_PCV201_5ms.RampUp) ,OTU(ControlLoop_PCV201_5ms.RampDown) ];
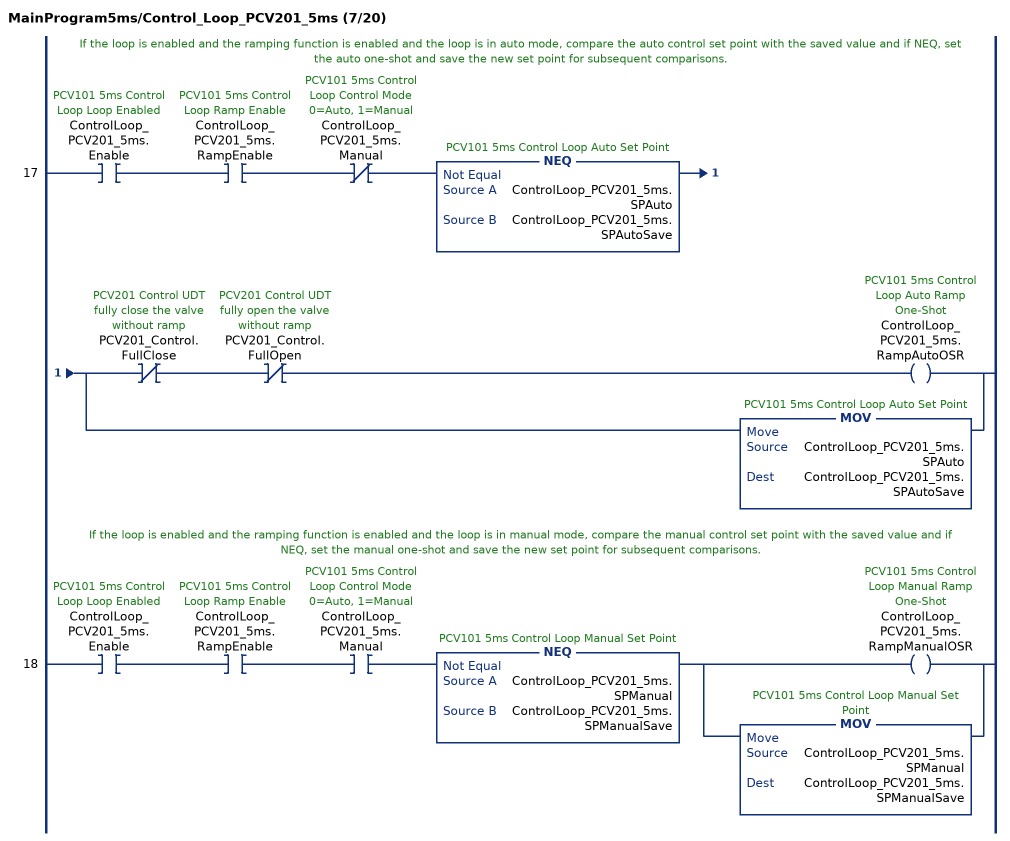
   // If the loop is enabled and the ramping function is enabled and the loop is in auto mode, compare the auto control set point with the saved value and if NEQ, set the auto one-shot and save the new set point for subsequent comparisons.
   17: XIC(ControlLoop_PCV201_5ms.Enable)XIC(ControlLoop_PCV201_5ms.RampEnable)XIO(ControlLoop_PCV201_5ms.Manual)NEQ(ControlLoop_PCV201_5ms.SPAuto,ControlLoop_PCV201_5ms.SPAutoSave)[XIO(PCV201_Control.FullClose) XIO(PCV201_Control.FullOpen) OTE(ControlLoop_PCV201_5ms.RampAutoOSR) ,MOV(ControlLoop_PCV201_5ms.SPAuto,ControlLoop_PCV201_5ms.SPAutoSave) ];
   // If the loop is enabled and the ramping function is enabled and the loop is in manual mode, compare the manual control set point with the saved value and if NEQ, set the manual one-shot and save the new set point for subsequent comparisons.
   18: XIC(ControlLoop_PCV201_5ms.Enable)XIC(ControlLoop_PCV201_5ms.RampEnable)XIC(ControlLoop_PCV201_5ms.Manual)NEQ(ControlLoop_PCV201_5ms.SPManual,ControlLoop_PCV201_5ms.SPManualSave)[OTE(ControlLoop_PCV201_5ms.RampManualOSR) ,MOV(ControlLoop_PCV201_5ms.SPManual,ControlLoop_PCV201_5ms.SPManualSave) ];
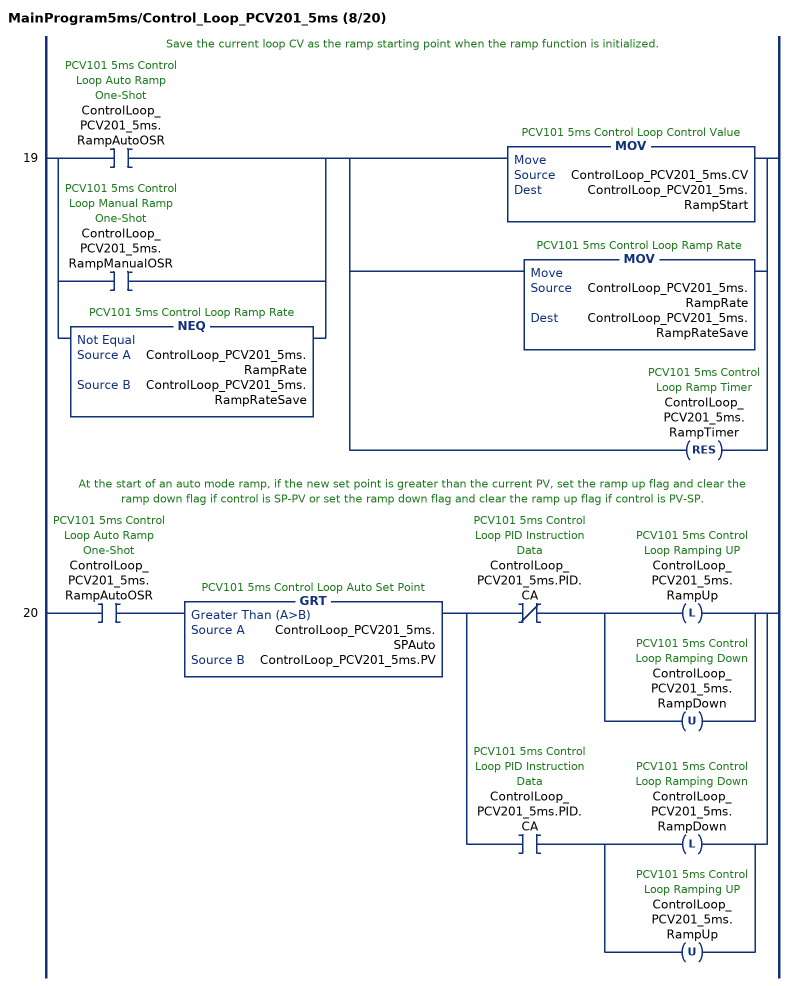
   // Save the current loop CV as the ramp starting point when the ramp function is initialized.
   19: [XIC(ControlLoop_PCV201_5ms.RampAutoOSR) ,XIC(ControlLoop_PCV201_5ms.RampManualOSR) ,NEQ(ControlLoop_PCV201_5ms.RampRate,ControlLoop_PCV201_5ms.RampRateSave) ][MOV(ControlLoop_PCV201_5ms.CV,ControlLoop_PCV201_5ms.RampStart) ,MOV(ControlLoop_PCV201_5ms.RampRate,ControlLoop_PCV201_5ms.RampRateSave) ,RES(ControlLoop_PCV201_5ms.RampTimer) ];
   // At the start of an auto mode ramp, if the new set point is greater than the current PV, set the ramp up flag and clear the ramp down flag if control is SP-PV or set the ramp down flag and clear the ramp up flag if control is PV-SP.
   20: XIC(ControlLoop_PCV201_5ms.RampAutoOSR)GRT(ControlLoop_PCV201_5ms.SPAuto,ControlLoop_PCV201_5ms.PV)[XIO(ControlLoop_PCV201_5ms.PID.CA) [OTL(ControlLoop_PCV201_5ms.RampUp) ,OTU(ControlLoop_PCV201_5ms.RampDown) ] ,XIC(ControlLoop_PCV201_5ms.PID.CA) [OTL(ControlLoop_PCV201_5ms.RampDown) ,OTU(ControlLoop_PCV201_5ms.RampUp) ] ];
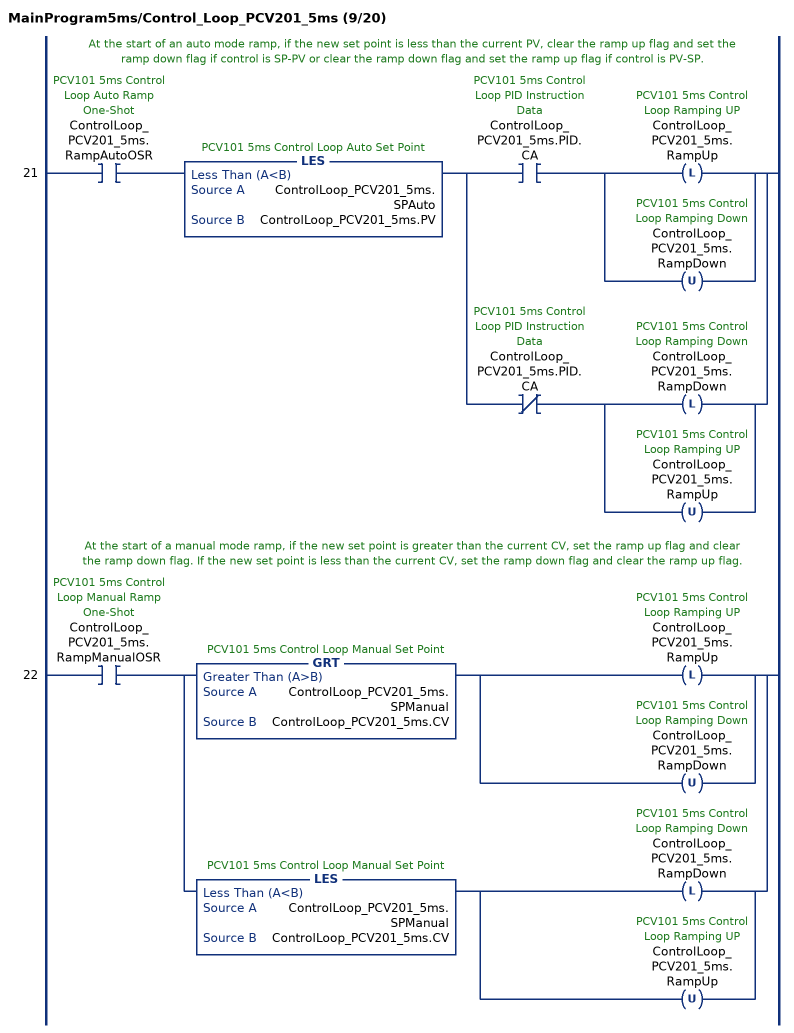
   // At the start of an auto mode ramp, if the new set point is less than the current PV, clear the ramp up flag and set the ramp down flag if control is SP-PV or clear the ramp down flag and set the ramp up flag if control is PV-SP.
   21: XIC(ControlLoop_PCV201_5ms.RampAutoOSR)LES(ControlLoop_PCV201_5ms.SPAuto,ControlLoop_PCV201_5ms.PV)[XIC(ControlLoop_PCV201_5ms.PID.CA) [OTL(ControlLoop_PCV201_5ms.RampUp) ,OTU(ControlLoop_PCV201_5ms.RampDown) ] ,XIO(ControlLoop_PCV201_5ms.PID.CA) [OTL(ControlLoop_PCV201_5ms.RampDown) ,OTU(ControlLoop_PCV201_5ms.RampUp) ] ];
   // At the start of a manual mode ramp, if the new set point is greater than the current CV, set the ramp up flag and clear the ramp down flag. If the new set point is less than the current CV, set the ramp down flag and clear the ramp up flag.
   22: XIC(ControlLoop_PCV201_5ms.RampManualOSR)[GRT(ControlLoop_PCV201_5ms.SPManual,ControlLoop_PCV201_5ms.CV) [OTL(ControlLoop_PCV201_5ms.RampUp) ,OTU(ControlLoop_PCV201_5ms.RampDown) ] ,LES(ControlLoop_PCV201_5ms.SPManual,ControlLoop_PCV201_5ms.CV) [OTL(ControlLoop_PCV201_5ms.RampDown) ,OTU(ControlLoop_PCV201_5ms.RampUp) ] ];
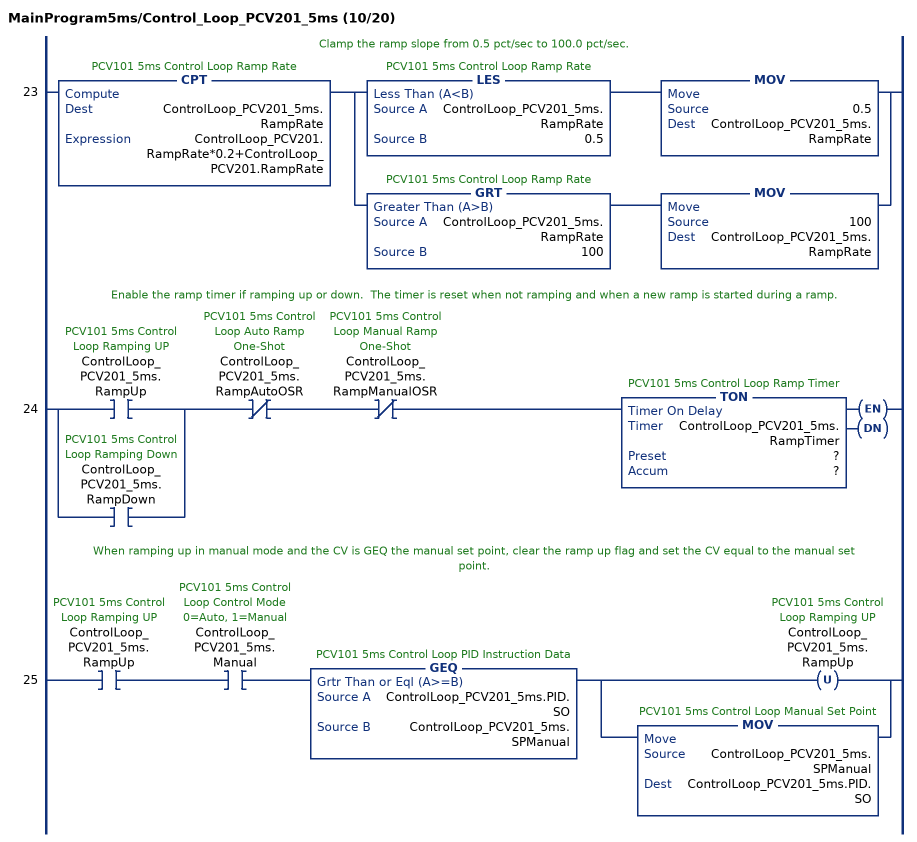
   // Clamp the ramp slope from 0.5 pct/sec to 100.0 pct/sec.
   23: CPT(ControlLoop_PCV201_5ms.RampRate,ControlLoop_PCV201.RampRate*0.2+ControlLoop_PCV201.RampRate)[LES(ControlLoop_PCV201_5ms.RampRate,0.5) MOV(0.5,ControlLoop_PCV201_5ms.RampRate) ,GRT(ControlLoop_PCV201_5ms.RampRate,100) MOV(100,ControlLoop_PCV201_5ms.RampRate) ];
   // Enable the ramp timer if ramping up or down.  The timer is reset when not ramping and when a new ramp is started during a ramp.
   24: [XIC(ControlLoop_PCV201_5ms.RampUp) ,XIC(ControlLoop_PCV201_5ms.RampDown) ]XIO(ControlLoop_PCV201_5ms.RampAutoOSR)XIO(ControlLoop_PCV201_5ms.RampManualOSR)TON(ControlLoop_PCV201_5ms.RampTimer,?,?);
   // When ramping up in manual mode and the CV is GEQ the manual set point, clear the ramp up flag and set the CV equal to the manual set point.
   25: XIC(ControlLoop_PCV201_5ms.RampUp)XIC(ControlLoop_PCV201_5ms.Manual)GEQ(ControlLoop_PCV201_5ms.PID.SO,ControlLoop_PCV201_5ms.SPManual)[OTU(ControlLoop_PCV201_5ms.RampUp) ,MOV(ControlLoop_PCV201_5ms.SPManual,ControlLoop_PCV201_5ms.PID.SO) ];
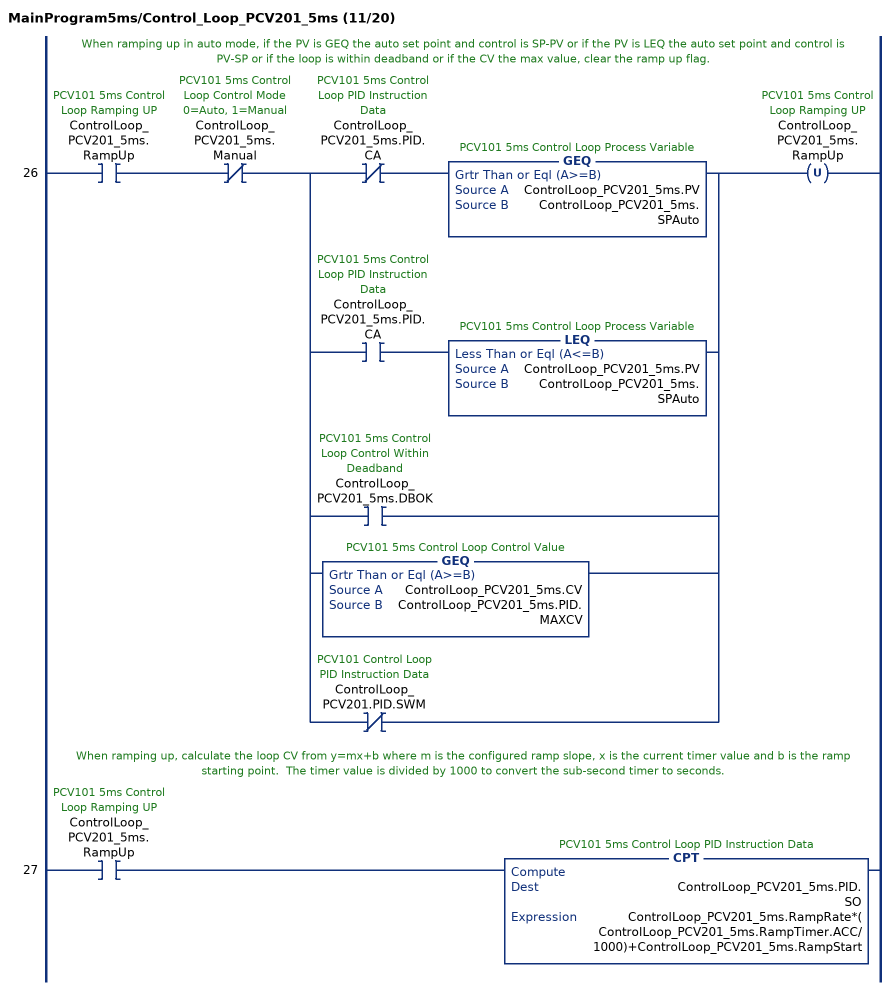
   // When ramping up in auto mode, if the PV is GEQ the auto set point and control is SP-PV or if the PV is LEQ the auto set point and control is PV-SP or if the loop is within deadband or if the CV the max value, clear the ramp up flag.
   26: XIC(ControlLoop_PCV201_5ms.RampUp)XIO(ControlLoop_PCV201_5ms.Manual)[XIO(ControlLoop_PCV201_5ms.PID.CA) GEQ(ControlLoop_PCV201_5ms.PV,ControlLoop_PCV201_5ms.SPAuto) ,XIC(ControlLoop_PCV201_5ms.PID.CA) LEQ(ControlLoop_PCV201_5ms.PV,ControlLoop_PCV201_5ms.SPAuto) ,XIC(ControlLoop_PCV201_5ms.DBOK) ,[GEQ(ControlLoop_PCV201_5ms.CV,ControlLoop_PCV201_5ms.PID.MAXCV) ,XIO(ControlLoop_PCV201.PID.SWM) ] ]OTU(ControlLoop_PCV201_5ms.RampUp);
   // When ramping up, calculate the loop CV from y=mx+b where m is the configured ramp slope, x is the current timer value and b is the ramp starting point.  The timer value is divided by 1000 to convert the sub-second timer to seconds.
   27: XIC(ControlLoop_PCV201_5ms.RampUp)CPT(ControlLoop_PCV201_5ms.PID.SO,ControlLoop_PCV201_5ms.RampRate*(ControlLoop_PCV201_5ms.RampTimer.ACC/1000)+ControlLoop_PCV201_5ms.RampStart);
